(* IEC 61131-3 sources: POMIRTS_lab3/AS/Library_2/ArTextSys, 3 files *)

(* ---- ArTextSys.typ ---- *)
TYPE
	ArTextSysLanguageCodeType : STRING[18]; (*String-type for language ID*)

	(*Enumeration for ArTextSysGetText-FUBs*)
	ArTextSysSearchModeEnum :
	(
		arTEXTSYS_SEARCH_FALLBACK_SUBST, (*with fallback-languages or substitute*)
		arTEXTSYS_SEARCH_LANGUAGE_ONLY, (*search for matching language only*)
		arTEXTSYS_SEARCH_FALLBACK	(*with fallback-searches, no substitute*)
	);

	(*argument-properties for formatter*)
	ArTextSysFormatArgumentType : STRUCT
		Datatype		: UINT;  (*type of argument; eg. IEC_DATATYPE_UDINT*)
		Data			: UDINT; (*pointer to Argument*)
		UnitNamespace	: UDINT; (*namespace of UnitID; default OPC-UA recommended*)
		UnitID			: UDINT;
	END_STRUCT;

	(*Internal type(s) for FUB-processing*)
	ArTextSysExec1InternalType : STRUCT
		i_serno : UINT;
		i_state : UINT;
		Result	: DINT;
	END_STRUCT;

	ArTextSysIter1InternalType : STRUCT
		i_base	: ArTextSysExec1InternalType;
		m_iter	: DINT; (*internal iterator; eg. ArTextSysGetNamespaceLanguages*)
	END_STRUCT;
END_TYPE

(* ---- ArTextSys.fun ---- *)
{REDUND_CONTEXT} {REDUND_UNREPLICABLE} FUNCTION_BLOCK ArTextSysGetSystemLanguage	(*determine preferred user-language*)
	VAR_INPUT
		Execute 		: BOOL; 			(*start on rising edge*)
	END_VAR
	VAR_OUTPUT
		Done			: BOOL; 			(*execution successful. FB finished*)
		Busy			: BOOL; 			(*FB is still active; needs call*)
		Error			: BOOL;
		StatusID		: DINT;
		LanguageCode	: ArTextSysLanguageCodeType;
	END_VAR
	VAR (*internals*)
		Internal : ArTextSysExec1InternalType;
	END_VAR
END_FUNCTION_BLOCK

{REDUND_CONTEXT} {REDUND_UNREPLICABLE} FUNCTION_BLOCK ArTextSysSetSystemLanguage	(*update preferred user-language*)
	VAR_INPUT
		Execute 		: BOOL;
		LanguageCode	: ArTextSysLanguageCodeType;
	END_VAR
	VAR_OUTPUT
		Done			: BOOL;
		Busy			: BOOL;
		Error			: BOOL; 			(*error occurred during operation*)
		StatusID		: DINT;
	END_VAR
	VAR (*internals*)
		Internal : ArTextSysExec1InternalType;
	END_VAR
END_FUNCTION_BLOCK

{REDUND_CONTEXT} {REDUND_UNREPLICABLE} FUNCTION_BLOCK ArTextSysGetNamespaceLanguages
	VAR_INPUT
		Execute 		: BOOL; 			(*start on rising edge*)
		Namespace		: UDINT;			(*string-pointer to namespace*)
		First			: BOOL; 			(*get first entry; or next*)
	END_VAR
	VAR_OUTPUT
		Done			: BOOL; 			(*execution successful. FB finished*)
		Busy			: BOOL; 			(*FB is still active; needs call*)
		Error			: BOOL; 			(*error occurred during operation*)
		StatusID		: DINT;
		LanguageCode	: ArTextSysLanguageCodeType;
		EndOfList		: BOOL; 			(*indicator for last found entry*)
	END_VAR
	VAR (*internals*)
		Internal : ArTextSysIter1InternalType;
	END_VAR
END_FUNCTION_BLOCK

{REDUND_CONTEXT} {REDUND_UNREPLICABLE} FUNCTION_BLOCK ArTextSysGetText
	VAR_INPUT
		Execute 		: BOOL;
		Namespace		: UDINT;			(*string-pointer to namespace*)
		TextID			: UDINT;			(*string-pointer to text-key*)
		LanguageCode	: ArTextSysLanguageCodeType;
		TextBufferSize	: UDINT;			(*size of result-buffer to get text*)
		TextBuffer		: UDINT;			(*pointer to text result-buffer*)
		SearchMode		: ArTextSysSearchModeEnum;
	END_VAR
	VAR_OUTPUT
		Done			: BOOL; 			(*execution successful. FB finished*)
		Busy			: BOOL; 			(*FB is still active; needs call*)
		Error			: BOOL; 			(*error occurred during operation*)
		StatusID		: DINT;
		TextSize		: UDINT;			(*Length of text in result-buffer*)
	END_VAR
	VAR (*internals*)
		Internal : ArTextSysExec1InternalType;
	END_VAR
END_FUNCTION_BLOCK

{REDUND_CONTEXT} {REDUND_UNREPLICABLE} FUNCTION_BLOCK ArTextSysFormatString
	VAR_INPUT
		Execute 		: BOOL;
		FormatString	: UDINT;			(*string-pointer to format-template*)
		ArgumentCount	: UINT; 			(*count of arguments in list*)
		ArgumentList	: ARRAY[0..9] OF ArTextSysFormatArgumentType;
		LanguageCode	: ArTextSysLanguageCodeType;
		MeasurementCode : UDINT;
		TextBufferSize	: UDINT;			(*size of result-buffer to get text*)
		TextBuffer		: UDINT;			(*pointer to result-buffer*)
	END_VAR
	VAR_OUTPUT
		Done			: BOOL; 			(*execution successful. FB finished*)
		Busy			: BOOL; 			(*FB is still active; needs call*)
		Error			: BOOL; 			(*error occurred during operation*)
		StatusID		: DINT;
		TextSize		: UDINT;			(*Length of text in result-buffer*)
	END_VAR
	VAR (*internals*)
		Internal : ArTextSysExec1InternalType;
	END_VAR
END_FUNCTION_BLOCK

{REDUND_CONTEXT} {REDUND_UNREPLICABLE} FUNCTION_BLOCK ArTextSysGetFormattedText
	VAR_INPUT
		Execute 		: BOOL;
		Namespace		: UDINT;			(*string-pointer to namespace*)
		TextID			: UDINT;			(*string-pointer to text-key*)
		ArgumentCount	: UINT; 			(*count of arguments in list*)
		ArgumentList	: ARRAY[0..9] OF ArTextSysFormatArgumentType;
		LanguageCode	: ArTextSysLanguageCodeType;
		MeasurementCode : UDINT;
		TextBufferSize	: UDINT;			(*size of result-buffer to get text*)
		TextBuffer		: UDINT;			(*pointer to result-buffer*)
		SearchMode		: ArTextSysSearchModeEnum;
	END_VAR
	VAR_OUTPUT
		Done			: BOOL; 			(*execution successful. FB finished*)
		Busy			: BOOL; 			(*FB is still active; needs call*)
		Error			: BOOL; 			(*error occurred during operation*)
		StatusID		: DINT;
		TextSize		: UDINT;			(*Length of text in result-buffer*)
	END_VAR
	VAR (*internals*)
		Internal : ArTextSysExec1InternalType;
	END_VAR
END_FUNCTION_BLOCK

(* ---- ArTextSys.var ---- *)
VAR CONSTANT
arTEXTSYS_ERR_OUT_OF_MEMORY 	: UDINT := 16#C030_280A;	(*fatal error: out of memory*)
arTEXTSYS_ERR_INVALID_ARG		: UDINT := 16#8030_280B;	(*provided argument is invalid*)
arTEXTSYS_ERR_FAILED			: UDINT := 16#8030_280C;	(*internal operation failure*)
arTEXTSYS_ERR_ACCESS_DENIED 	: UDINT := 16#8030_280D;	(*resource-access denied*)
arTEXTSYS_ERR_INVALID_HANDLE	: UDINT := 16#8030_280E;	(*invalid handle detected*)

arTEXTSYS_ERR_CANT_OPEN_TEXTDB	: UDINT := 16#8030_2811;	(*opening of text-db failed*)
arTEXTSYS_INF_ALREADY_OPENED	: DINT	:= 16#4030_2812;	(*text-db is open and ready*)
arTEXTSYS_ERR_TEXTDB_SCHEMA 	: UDINT := 16#8030_2813;	(*unrecognised text-db schema or structure*)
arTEXTSYS_ERR_TEXTDB_READER 	: UDINT := 16#8030_2814;	(*read of open text-db failed*)
arTEXTSYS_ERR_TEXTDB_INTERNAL	: UDINT := 16#8030_2815;	(*other kind of text-db error*)
arTEXTSYS_INF_NOT_SET_DURABLE	: DINT	:= 16#4030_2816;	(*configuration-change is not durable*)

arTEXTSYS_ERR_NO_TEXT_FOUND 	: UDINT := 16#8030_2818;	(*no requested text found*)
arTEXTSYS_INF_LANGUAGE_DIFFERS	: DINT	:= 16#4030_281A;	(*text-language differs; not in requested language*)
arTEXTSYS_INF_SUBSTITUTE_TEXT	: DINT	:= 16#4030_281B;	(*no text found, but substitute-text provided*)
arTEXTSYS_ERR_NOT_EXISTS		: UDINT := 16#8030_281C;	(*record not found; doesn't exist*)
arTEXTSYS_ERR_END_REACHED		: UDINT := 16#8030_281D;	(*no further suitable entry found*)
END_VAR
